// TIA Portal V17 export
FUNCTION_BLOCK "FB_T06_Commente"   // FB106, LAD
TITLE = Surveillance niveau
{ S7_Optimized_Access := 'TRUE' }
// Bloc de test : commentaires, valeurs initiales, constante.
// stored: IsIECCheckEnabled false, MemoryReserve 100, SetENOAutomatically false
   VAR_INPUT
      Niveau : Int := 0;   // Niveau cuve (0..1000)
   END_VAR
   VAR_OUTPUT
      Alarme : Bool := false;   // Alarme niveau haut
   END_VAR
   VAR
      Actif : Bool := true;   // Surveillance active
      Nb_Alarmes : Int := 0;   // Compteur d'alarmes
   END_VAR
   VAR_TEMP
      Tmp : Bool;   // Variable temporaire
   END_VAR
   VAR CONSTANT
      SEUIL_HAUT : Int := 800;   // Seuil de déclenchement
   END_VAR
BEGIN

REGION Network 1: Alarme niveau haut
   // Déclenche l'alarme quand le niveau atteint le seuil.
   // Seuil défini par la constante SEUIL_HAUT.
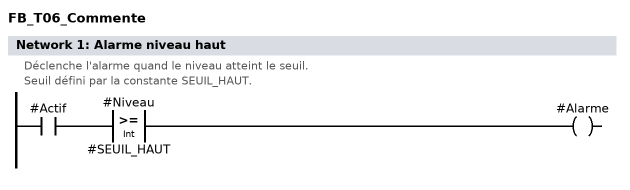
   #Alarme := #Actif AND (#Niveau >= #SEUIL_HAUT);
END_REGION
END_FUNCTION_BLOCK
